(* IEC 61131-3 sources: Lasal-MCP/examples/SampleSource/LASALScreenAdvancedSolution/LASALScreenAdvancedSolution/LASALScreenAdvacnedSolution/Stations/Terminal/HMI/Class/MyCarousel, 1 file *)

(* ---- MyCarousel.st ---- *)
#define MAX_ITEMS 20

//***** Parameters for Carousel *****
#define HORIZONTAL_DRAW_ORDER_CARO FALSE
#define INFINITE_CARO FALSE
#define ELEMENT_GAP_CARO 5
#define FRAMEWORK_NEW_AGE_DARK 81 // ID in LSE
#define VERTICAL_SCROLL_BAR TRUE

(*!
<Class
	Name               = "MyCarousel"
	Revision           = "0.0"
	RealtimeTask       = "false"
	CyclicTask         = "false"
	BackgroundTask     = "false"
	Sigmatek           = "false"
	OSInterface        = "false"
	HighPriority       = "false"
	Automatic          = "false"
	UpdateMode         = "Prescan"
	SharedCommandTable = "true"
	Objectsize         = "(538,120)">
	<Channels>
		<Server Name="LasalObjectName" Class="StringInternal" Visualized="true" Remotely="true" Initialize="true" WriteProtected="false" Retentive="false"/>
		<Server Name="LSEObjectName" Class="StringInternal" Visualized="true" Remotely="true" Initialize="true" WriteProtected="false" Retentive="false"/>
		<Server Name="ShowActive" Visualized="true" Initialize="false" WriteProtected="false" Retentive="false"/>
		<Server Name="xy1x" Visualized="false" Initialize="true" WriteProtected="true" Retentive="false"/>
		<Server Name="xy1y" Visualized="false" Initialize="true" WriteProtected="true" Retentive="false"/>
		<Server Name="xy2x" Visualized="false" Initialize="true" WriteProtected="true" Retentive="false"/>
		<Server Name="xy2y" Visualized="false" Initialize="true" WriteProtected="true" Retentive="false"/>
		<Client Name="LasalObjName" Required="true" Internal="true"/>
		<Client Name="LSEObjName" Required="true" Internal="true"/>
		<Client Name="SigCLib" Required="false" Internal="false"/>
	</Channels>
	<Network Name="MyCarousel">
		<!-- List of Components in this network -->
		<Components>
			<Object
				Name       = "_base"
				Class      = "_Screen"
				Position   = "(218,120)"
				Visualized = "true"
				Remotely   = "true">
				<Channels>
					<Server Name="Screen"/>
					<Client Name="ImA"/>
					<Client Name="Lse"/>
					<Client Name="No"/>
				</Channels>
			</Object>
			<Object
				Name       = "LasalObjName"
				Class      = "StringRAM"
				Position   = "(210,480)"
				Visualized = "true"
				Remotely   = "true">
				<Channels>
					<Server Name="Data" Value="MyValues"/>
					<Client Name="SingleRealloc" Value="1"/>
					<Client Name="UseFile"/>
				</Channels>
			</Object>
			<Object
				Name       = "LSEObjName"
				Class      = "StringRAM"
				Position   = "(210,720)"
				Visualized = "true"
				Remotely   = "true">
				<Channels>
					<Server Name="Data" Value="Value"/>
					<Client Name="SingleRealloc" Value="1"/>
					<Client Name="UseFile"/>
				</Channels>
			</Object>
		</Components>
		<Comments>
		</Comments>
		<!-- List of Connections in this network -->
		<Connections>
			<Connection Source="this.Screen" Destination="_base.Screen" Vertices="(878,210),(518,210),"/>
			<Connection Source="_base.Lse" Destination="this.Lse" Vertices="(218,210),(38,210),"/>
			<Connection Source="_base.No" Destination="this.No" Vertices="(218,270),(38,270),"/>
			<Connection Source="_base.ImA" Destination="this.ImA" Vertices="(218,330),(38,330),"/>
			<Connection Source="this.LasalObjName" Destination="LasalObjName.Data"/>
			<Connection Source="this.LSEObjName" Destination="LSEObjName.Data"/>
			<Connection Source="this.LasalObjectName" Destination="LasalObjName.Data" Vertices="(878,390),(706,570),"/>
			<Connection Source="this.LSEObjectName" Destination="LSEObjName.Data" Vertices="(878,450),(706,810),"/>
		</Connections>
		<!-- Headerfiles -->
		<Options>
		</Options>
	</Network>
</Class>
*)
#pragma using _Screen

MyCarousel : CLASS
: _Screen
  //Servers:
	LasalObjectName 	: SvrChCmd_UDINT;
	LSEObjectName 	: SvrChCmd_UDINT;
	xy1x 	: SvrCh_DINT;
	xy1y 	: SvrCh_DINT;
	xy2x 	: SvrCh_DINT;
	xy2y 	: SvrCh_DINT;
	ShowActive 	: SvrCh_DINT;
  //Clients:
	LasalObjName 	: CltChCmd_StringRAM;
	LSEObjName 	: CltChCmd_StringRAM;
	SigCLib 	: CltChCmd_SigCLib;
  //Variables:
		localLasalObjName : ARRAY [0..255] OF CHAR;

		localLSEObjName : ARRAY [0..255] OF CHAR;

		intError 	: DINT;
		myCaroItems : ARRAY [1..MAX_ITEMS] OF _CAROITEM;

		carousel 	: DINT;
		noOfCarouselItems 	: UDINT;
		pError 	: ^CHAR;
  //Functions:

	FUNCTION VIRTUAL GLOBAL Init;

	FUNCTION VIRTUAL GLOBAL S_Start
		VAR_INPUT
			pic 	: ^void;
			firsttime 	: BOOL;
		END_VAR;

	FUNCTION VIRTUAL GLOBAL InitObjNames;

	FUNCTION PlaceCarousel
		VAR_INPUT
			pPic 	: ^void;
			pLasalObjName 	: ^CHAR;
			pLSEObjName 	: ^CHAR;
			Room 	: _ROOM;
			CaroItemsCount 	: UDINT;
			VarNoPos 	: UDINT;
		END_VAR
		VAR_OUTPUT
			Retcode 	: DINT;
		END_VAR;

	FUNCTION AddItem
		VAR_INPUT
			ObjNo 	: UDINT;
			LasalObjNo 	: UDINT;
			CarItemNo 	: UDINT;
		END_VAR
		VAR_OUTPUT
			Retcode 	: DINT;
		END_VAR;

	FUNCTION VIRTUAL GLOBAL LasalObjectName::Read
		VAR_OUTPUT
			output (EAX) 	: UDINT;
		END_VAR;

	FUNCTION VIRTUAL GLOBAL LasalObjectName::Write
		VAR_INPUT
			input (EAX) 	: UDINT;
		END_VAR
		VAR_OUTPUT
			result (EAX) 	: UDINT;
		END_VAR;

	FUNCTION VIRTUAL GLOBAL LSEObjectName::Read
		VAR_OUTPUT
			output (EAX) 	: UDINT;
		END_VAR;

	FUNCTION VIRTUAL GLOBAL LSEObjectName::Write
		VAR_INPUT
			input (EAX) 	: UDINT;
		END_VAR
		VAR_OUTPUT
			result (EAX) 	: UDINT;
		END_VAR;

	FUNCTION VIRTUAL GLOBAL ShowActive::Write
		VAR_INPUT
			input (EAX) 	: DINT;
		END_VAR
		VAR_OUTPUT
			result (EAX) 	: DINT;
		END_VAR;
  //Tables:
	FUNCTION @STD
		VAR_OUTPUT
			ret_code	: CONFSTATES;
		END_VAR;
	FUNCTION GLOBAL TAB @CT_;
END_CLASS;

#pragma using StringRAM
#pragma usingLtd SigCLib

#pragma usingltd MyValues

FUNCTION VIRTUAL GLOBAL MyCarousel::Init
VAR
  number : USINT;
END_VAR

  _Screen::Init(); // call method of base

  if (_FirstScan = TRUE) then
    InitObjNames();

    for number := 1 to (MAX_ITEMS) do
      init_CAROITEM(p:= #myCaroItems[number]);
      init_VARLABEL(p0:= #myCaroItems[number].loader);
    end_for;

  end_if;

END_FUNCTION

FUNCTION VIRTUAL GLOBAL MyCarousel::InitObjNames
VAR
	strLength : UDINT;
END_VAR

  // get object name from values
  strLength := LasalObjName.GetLength();

  LasalObjName.GetDataAt(pData:= #localLasalObjName[0],
                         udSize:= strLength,
                         udAt:= 0);

  localLasalObjName[strLength] := 0;

  // get object name from screen
  strLength := LSEObjName.GetLength();

  LSEObjName.GetDataAt(pData:= #localLSEObjName[0],
                       udSize:= strLength,
                       udAt:= 0);

  localLSEObjName[strLength] := 0;

  carousel := -1;

END_FUNCTION

FUNCTION VIRTUAL GLOBAL MyCarousel::S_Start
	VAR_INPUT
		pic 	: ^void;
		firsttime 	: BOOL;
	END_VAR
  VAR
  	room : _ROOM;
  END_VAR

  _Screen::S_Start(pic:= pic, firsttime:= firsttime);

  if (firsttime = TRUE) then

    room.xy1.x := to_int(xy1x);
    room.xy1.y := to_int(xy1y);
    room.xy2.x := to_int(xy2x);
    room.xy2.y := to_int(xy2y);

    intError := PlaceCarousel(pPic:= pic,
                              pLasalObjName:= #localLasalObjName[0],
                              pLSEObjName:= #localLSEObjName[0],
                              Room:= room,
                              CaroItemsCount:= MAX_ITEMS,
                              VarNoPos:= 20);
  end_if;

END_FUNCTION

FUNCTION MyCarousel::PlaceCarousel
	VAR_INPUT
		pPic 	: ^void;
		pLasalObjName 	: ^CHAR;
		pLSEObjName 	: ^CHAR;
		Room 	: _ROOM;
		CaroItemsCount 	: UDINT;
		VarNoPos 	: UDINT;
	END_VAR
	VAR_OUTPUT
		Retcode 	: DINT;
	END_VAR
  VAR
    index         : UDINT;
    caroItem      : UDINT;
    objectName    : ARRAY[0..255]of CHAR;
    objectNumber  : ARRAY[0..255]of CHAR;
    objectNo      : UDINT;
    lasalObjectNo : UDINT;
    varinfo       : _VARINFO;
    retGetVarInfo : BOOL;
  END_VAR

  Retcode := 0;

  // check for valid pointers
  if ((pPic = NIL) | (pLasalObjName = NIL) | (pLSEObjName = NIL)) then
    Retcode := -1; // invalid pointers
    return;
  end_if;

  objectNo := get_no_by_label(p0:= pLSEObjName,
                              x1:= OBJLST,
                              x2:= 0);

  if (objectNo = DEFSCOPE) then
    Retcode := -2; // invalid LSE objectname
    return;
  end_if;

  if (CaroItemsCount > MAX_ITEMS) then
    Retcode := -3; // to much items
    return;
  end_if;

  noOfCarouselItems := 0;
  caroItem := 1;

  for index := 1 to (CaroItemsCount) do

    pError := SigCLib.StrCpy(dst0:= #objectName[0],
                             src0:= pLasalObjName);

    if (pError <> #objectName[0]) then
      Retcode := -4;
      return;
    end_if;

    objectNumber[0] := 0;

    pError := SigCLib.IToA(val:= to_dint(index),
                           dst:= #objectNumber[0],
                           base:= 10);

    if (pError <> #objectNumber[0]) then
      Retcode := -5;
      return;
    end_if;

    pError := SigCLib.StrCat(ps1:= #objectName[0],
                             ps2:= #objectNumber[0]);

    if (pError <> #objectName[0]) then
      Retcode := -6;
      return;
    end_if;

    lasalObjectNo := VarList_GetVarNoStation(p0:= #objectName[0],
                                             station:= 255);

    if (lasalObjectNo = DEFSCOPE) then
      Retcode := -7; // invalid objectname / no
      return;
    end_if;

    retGetVarInfo := VarList_GetVarInfo(p0:= #varinfo,
                                        x1:= lasalObjectNo);

    if (retGetVarInfo = FALSE) then
      Retcode := -8; // no var info found
      return;
    end_if;

    if (varinfo.lasalid.id = 0) then
      Retcode := -9; // wrong lasal ID
      return;
    end_if;

    if (ShowActive = 1) then

      if (varinfo.lasalid.id$^MyValues^.Active.Read()) then

        Retcode := AddItem(ObjNo:= objectNo,
                           LasalObjNo:= lasalObjectNo,
                           CarItemNo:= caroItem);

        caroItem += 1;
        noOfCarouselItems += 1;

      end_if;

    else
      Retcode := AddItem(ObjNo:= objectNo,
                         LasalObjNo:= lasalObjectNo,
                         CarItemNo:= caroItem);

      caroItem += 1;
      noOfCarouselItems += 1;

    end_if;

  end_for;

  for index := caroItem to (CaroItemsCount) do
    myCaroItems[index].ObjNo := 0;
    init_VARLABEL(p0:= #myCaroItems[index].loader);
  end_for;

  carousel := add_carousel(mp:= pPic$^_MY_PICTURE,
                           room:= #Room,
                           cino:= to_uint(noOfCarouselItems),
                           ci:= #myCaroItems[1],
                           varno_pos:= DEFSCOPE,
                           horizontal:= HORIZONTAL_DRAW_ORDER_CARO,
                           infinite:= INFINITE_CARO,
                           _dx:= ELEMENT_GAP_CARO);

  #pragma warning(disable:69);
  if (VERTICAL_SCROLL_BAR) then
  #pragma warning(default:69);

    add_carousel_scrollbar(mp:= pPic$^_MY_PICTURE,
                           cno:= carousel,
                           frame:= FRAMEWORK_NEW_AGE_DARK,
                           col_back:= LSE_COLOR252,
                           col_front:= LSE_color246,
                           col_symbol:= LSE_COLOR255,
                           col_topleft:= INVISIBLE,
                           col_bottomright:= INVISIBLE);
  end_if;

  Retcode := 1;

END_FUNCTION

FUNCTION MyCarousel::AddItem
	VAR_INPUT
		ObjNo 	: UDINT;
		LasalObjNo 	: UDINT;
		CarItemNo 	: UDINT;
	END_VAR
	VAR_OUTPUT
		Retcode 	: DINT;
	END_VAR
  VAR
  	result : _RESULT;
    variable : _VARIABLE;
  END_VAR

  Retcode := 0;

  myCaroItems[CarItemNo].ObjNo := TO_UINT(ObjNo);

  #pragma warning(disable:74);
  myCaroItems[CarItemNo].loader.no := 1;
  myCaroItems[CarItemNo].loader.info[0].state := VAR_VAL;
  myCaroItems[CarItemNo].loader.info[0].value := TO_DINT(LasalObjNo);
  #pragma warning(default:74);

  if (VarList_GetSystemData(p0:= #result,
                            p1:= #variable,
                            p2:= #myCaroItems[CarItemNo].loader,
                            x3:= true) = TRUE) then
    Retcode := -7;
    return;
  end_if;

END_FUNCTION

FUNCTION VIRTUAL GLOBAL MyCarousel::ShowActive::Write
	VAR_INPUT
		input (EAX) 	: DINT;
	END_VAR
	VAR_OUTPUT
		result (EAX) 	: DINT;
	END_VAR

	ShowActive := input;
	result := ShowActive;

  InsertCmd(x0:= CMD_NEWPICTURE, x1:= to_DINT(No), x2:= 0);

END_FUNCTION

FUNCTION VIRTUAL GLOBAL MyCarousel::LasalObjectName::Read
	VAR_OUTPUT
		output (EAX) 	: UDINT;
	END_VAR

	LasalObjectName := LasalObjName.Data.Read();
	output := LasalObjectName;

END_FUNCTION

FUNCTION VIRTUAL GLOBAL MyCarousel::LasalObjectName::Write
	VAR_INPUT
		input (EAX) 	: UDINT;
	END_VAR
	VAR_OUTPUT
		result (EAX) 	: UDINT;
	END_VAR

	LasalObjectName := input;
	result := (LasalObjName.Data.Write(LasalObjectName))$UDINT;

END_FUNCTION

FUNCTION VIRTUAL GLOBAL MyCarousel::LSEObjectName::Read
	VAR_OUTPUT
		output (EAX) 	: UDINT;
	END_VAR

	LSEObjectName := LSEObjName.Data.Read();
	output := LSEObjectName;

END_FUNCTION

FUNCTION VIRTUAL GLOBAL MyCarousel::LSEObjectName::Write
	VAR_INPUT
		input (EAX) 	: UDINT;
	END_VAR
	VAR_OUTPUT
		result (EAX) 	: UDINT;
	END_VAR

	LSEObjectName := input;
	result := (LSEObjName.Data.Write(LSEObjectName))$UDINT;

END_FUNCTION
